(* IEC 61131-3 sources: nautilus/logix/writer/testdata/conformance/yardstick/lib, 1 file *)

(* ---- types.st ---- *)
TYPE
  LineStatus : STRUCT
    Mode  : DINT;
    Alarm : BOOL;
  END_STRUCT;
END_TYPE
